Staubli VAL3: frameItem.dtx

public string sName
public frame fFrame = {fatherId=world[0]}
public pointRx pPointRx[3]
  [0] = {fatherId=world[0]}
  [1] = {fatherId=world[0]}
  [2] = {fatherId=world[0]}
